FUNCTION_BLOCK FB_TerminalDiagnosis
VAR_INPUT
	stTerminalState				:ST_TerminalState;
END_VAR
VAR_OUTPUT
	bTerminalOK					:BOOL;
	sTerminalStatus				:STRING;
END_VAR
VAR

	sStateStatusAll				:STRING(255);
	sState						:STRING;
	sWorkingState				:STRING;
	tonTerminalNOK				:TON;
END_VAR
VAR CONSTANT
	tTerminalNOKDelay				:TIME := t#2s;
END_VAR

(*This Function returns the State of the Device. Either one of the States INIT, PREOP, OP, BOOTSTRAP or SAFE-OP is returned. stState is given the Value of the Function. *)
sState:= F_StateReturn(state:= stTerminalState.unInfoState);

(*All other Errors that can occur concerning the State of the Device*)
(*Because theoratically all the other errors could occur all together, CONCAT is done to show them all in one view box.*)
IF stTerminalState.unInfoState.4
THEN
	sStateStatusAll:= 'Slave signals error. ';
ELSE
	sStateStatusAll:= '';
END_IF

IF stTerminalState.unInfoState.5
THEN
	sStateStatusAll:= CONCAT( sStateStatusAll, 'Invalid vendorID. ');
ELSE
	sStateStatusAll:= CONCAT( sStateStatusAll, '');
END_IF

IF stTerminalState.unInfoState.6
THEN
	sStateStatusAll:= CONCAT( sStateStatusAll, 'Initialization error occurred. ');
ELSE
	sStateStatusAll:= CONCAT( sStateStatusAll, '');
END_IF

IF stTerminalState.unInfoState.7
THEN
	sStateStatusAll:= CONCAT( sStateStatusAll, 'Slave disabled. ');
ELSE
	sStateStatusAll:= CONCAT( sStateStatusAll, '');
END_IF

IF stTerminalState.unInfoState.8
THEN
	sStateStatusAll:= CONCAT( sStateStatusAll, 'Slave not present. ');
ELSE
	sStateStatusAll:= CONCAT( sStateStatusAll, '');
END_IF

IF stTerminalState.unInfoState.9
THEN
	sStateStatusAll:= CONCAT( sStateStatusAll, 'Slave signals link error. ');
ELSE
	sStateStatusAll:= CONCAT( sStateStatusAll, '');
END_IF

IF stTerminalState.unInfoState.10
THEN
	sStateStatusAll:= CONCAT( sStateStatusAll, 'Slave signals missing link. ');
ELSE
	sStateStatusAll:= CONCAT( sStateStatusAll, '');
END_IF

IF stTerminalState.unInfoState.11
THEN
	sStateStatusAll:= CONCAT( sStateStatusAll, 'Slave signals unexpected link. ');
ELSE
	sStateStatusAll:= CONCAT( sStateStatusAll, '');
END_IF

IF stTerminalState.unInfoState.12
THEN
	sStateStatusAll:= CONCAT( sStateStatusAll,  'Communication port A. ');
ELSE
	sStateStatusAll:= CONCAT( sStateStatusAll, '');
END_IF

IF stTerminalState.unInfoState.13
THEN
	sStateStatusAll:= CONCAT( sStateStatusAll, 'Communication port B. ');
ELSE
	sStateStatusAll:= CONCAT( sStateStatusAll, '');
END_IF

IF stTerminalState.unInfoState.14
THEN
	sStateStatusAll:= CONCAT( sStateStatusAll, 'Communication port C. ');
ELSE
	sStateStatusAll:= CONCAT( sStateStatusAll, '');
END_IF

IF stTerminalState.unInfoState.15
THEN
	sStateStatusAll:= CONCAT( sStateStatusAll,  'Communication port D. ');
ELSE
	sStateStatusAll:= CONCAT( sStateStatusAll, '');
END_IF

(*If none of the other errors occur, the text of the view box is 'None'.*)
IF sStateStatusAll= ''
THEN
	sStateStatusAll:= 'No error';
END_IF

(*The colour and text of the view box WcState is adjusted.*)
IF stTerminalState.bWcState = 0
THEN
	sWorkingState:= 'Working State OK ';
ELSE
	sWorkingState:= 'Working State NOT OK ';
END_IF

(*General Status Information*)
bTerminalOK:= TRUE;
sTerminalStatus:= 'Terminal OK ';

IF stTerminalState.bWcState <> 0
     OR sStateStatusAll <> 'No error'
THEN
	tonTerminalNOK(IN := TRUE, PT := tTerminalNOKDelay);
	IF tonTerminalNOK.Q
	THEN
		bTerminalOK:= FALSE;
		sTerminalStatus:= 'Terminal Error ';
	ELSE
		sTerminalStatus:= 'Waiting for status.';
	END_IF
END_IF

END_FUNCTION_BLOCK

(* stored: Version 1.1.0.1, ProductVersion 3.1.4024.15
   POU FB_TerminalDiagnosis: Id {d76ebce7-4726-47a6-a477-2d5273d32cae}, SpecialFunc None *)
